Fanuc KAREL source: KD00070.KL

PROGRAM KD00070
%NOLOCKGROUP
VAR
  I: INTEGER
  J: INTEGER
  B: BOOLEAN
  R: REAL
  S: STRING[80]
BEGIN
  CONDITION[1]:
  WHEN DIN[1] = ON DO
    STOP
  ENDCONDITION
END KD00070
